TYPE ST_Tapahtumaloki :
STRUCT
	nID:				LINT;
	tAikaleima:			DATE_AND_TIME;
	sTapahtuma:			STRING(50);
	sKuvaus:			STRING(255);

	
END_STRUCT
END_TYPE

(* stored: Version 1.1.0.1
   DUT ST_Tapahtumaloki: Id {51130b9f-bee3-41a2-bf83-5378b8e48a55} *)
